FUNCTION fun_LrealToString : STRING
VAR_INPUT
	iDigits	: INT:=2;
	fVar	: LREAL;
END_VAR
VAR
	iDigitsLocal: INT;

	fTemp: LREAL;
	fMult: LREAL;
	
	fbFormat: FB_FormatString;	

END_VAR

IF iDigits<0 THEN;
	iDigitsLocal:=0;
ELSIF iDigits>6 THEN;
	iDigitsLocal:=6; 
ELSE
	iDigitsLocal:=iDigits;	
END_IF

// this vertion solve the case then the result is 2.0-e2 instade of 0.02
CASE iDigitsLocal OF
	0:;fbFormat(sFormat:='%.0f' ,arg1:=F_LREAL(fVar),sOut=>fun_LrealToString);
	1:;fbFormat(sFormat:='%.1f' ,arg1:=F_LREAL(fVar),sOut=>fun_LrealToString);
	2:;fbFormat(sFormat:='%.2f' ,arg1:=F_LREAL(fVar),sOut=>fun_LrealToString);
	3:;fbFormat(sFormat:='%.3f' ,arg1:=F_LREAL(fVar),sOut=>fun_LrealToString);
	4:;fbFormat(sFormat:='%.4f' ,arg1:=F_LREAL(fVar),sOut=>fun_LrealToString);
	5:;fbFormat(sFormat:='%.5f' ,arg1:=F_LREAL(fVar),sOut=>fun_LrealToString);
	6:;fbFormat(sFormat:='%.6f' ,arg1:=F_LREAL(fVar),sOut=>fun_LrealToString);
END_CASE

(* OLD Version
CASE iDigitsLocal OF
	0:;fMult:=1;
	1:;fMult:=10;
	2:;fMult:=100;
	3:;fMult:=1000;
	4:;fMult:=10000;
	5:;fMult:=100000;
	6:;fMult:=1000000;
END_CASE

fTemp:=TRUNC(fVar*fMult);
IF iDigitsLocal=0 THEN;
	fun_LrealToString:=DINT_TO_STRING(TRUNC(fVar));
ELSE;
	fun_LrealToString:=LREAL_TO_STRING(fTemp/fMult);	
END_IF
*)

END_FUNCTION

(* stored: Version 1.1.0.1, ProductVersion 3.1.4024.12
   POU fun_LrealToString: Id {7566430a-b270-46a7-aa63-4244670fe50f}, SpecialFunc None *)
